Fanuc KAREL source: KT00900.KL

PROGRAM KT00900
%NOLOCKGROUP
VAR
  P1: XYZWPREXT
  P2: XYZWPREXT
  OUT: BOOLEAN
BEGIN
  P1.X = 1.0
  P2.Y = 2.0
  P1.X = 1.0
  P2.Y = 2.0
  OUT = J_IN_RANGE(P1)
END KT00900
